FUNCTION_BLOCK FB_MotionSystem
VAR
    fbXPlanarSystem   : FB_XPlanarSystem;
    fbXPlanarMover    : ARRAY[1..maxNumMover] OF FB_XPlanarMoverStandard;
    nStartupSequence  : UDINT;
    nStartingSequence : UDINT;
    nExecutingSequence : UDINT;
    nErrorStep         : UDINT;    // step where the error happened
    nErrorID           : UDINT;    // error code of the motion command
END_VAR

METHOD Cycle
VAR
    i : UDINT;
END_VAR
// Call every PLC cycle: updates the XPlanar system and the movers.
fbXPlanarSystem.Cycle();
FOR i := 1 TO moverCount DO
    fbXPlanarMover[i].Cycle();
END_FOR
END_METHOD

METHOD Execute6DoF : BOOL
VAR_INPUT
    bReset : BOOL;
END_VAR
VAR_INST
    stStartPos   : PositionXYC;
    stCenterPos  : PositionXYC;
    stRotOptions : ST_MoveCOptions;
END_VAR
// One 6 DoF sequence with mover 1. TRUE when finished. Stops in step 900 on error.
IF bReset THEN
    Execute6DoF := FALSE;
    nExecutingSequence := 0;
    nErrorStep := 0;
    nErrorID := 0;
END_IF

CASE nExecutingSequence OF
    // store the start position
    0:  stStartPos.SetValuesXYC(fbXPlanarMover[1].P_ActPosition.x,
                                fbXPlanarMover[1].P_ActPosition.y,
                                fbXPlanarMover[1].P_ActPosition.c);
        stCenterPos.SetValuesXYC(480, 360, 0);
        stRotOptions.additionalTurns := 0;
        stRotOptions.direction := Tc3_Mc3PlanarMotion.MC_Direction.mcDirectionNonModulo;
        IF NOT bReset THEN
            nExecutingSequence := 10;
        END_IF

    // drive to the table centre
    10: fbXPlanarMover[1].MoveToPosition('To center', stCenterPos, 500, 1250, 1250, 12500);
        nExecutingSequence := 11;
    11: IF fbXPlanarMover[1].P_MoveToPosition.Done THEN
            nExecutingSequence := 20;
        ELSIF fbXPlanarMover[1].P_MoveToPosition.Error THEN
            nErrorStep := nExecutingSequence;
            nErrorID := fbXPlanarMover[1].P_MoveToPosition.ErrorID;
            nExecutingSequence := 900;
        END_IF

    // lift Z to 4 mm
    20: fbXPlanarMover[1].MoveZ('Z up', 4, 20, 100, 100, 1000);
        nExecutingSequence := 21;
    21: IF fbXPlanarMover[1].P_MoveZ.Done THEN
            nExecutingSequence := 30;
        ELSIF fbXPlanarMover[1].P_MoveZ.Error THEN
            nErrorStep := nExecutingSequence;
            nErrorID := fbXPlanarMover[1].P_MoveZ.ErrorID;
            nExecutingSequence := 900;
        END_IF

    // rotate C +90 deg
    30: fbXPlanarMover[1].MoveC('C +90', 90, 720, 1800, 1800, 9000, stRotOptions);
        nExecutingSequence := 31;
    31: IF fbXPlanarMover[1].P_MoveC.Done THEN
            nExecutingSequence := 50;
        ELSIF fbXPlanarMover[1].P_MoveC.Error THEN
            nErrorStep := nExecutingSequence;
            nErrorID := fbXPlanarMover[1].P_MoveC.ErrorID;
            nExecutingSequence := 900;
        END_IF

	// lower Z
	40: fbXPlanarMover[1].MoveZ('Z down', 2, 20, 100, 100, 1000);
        nExecutingSequence := 41;
    41: IF fbXPlanarMover[1].P_MoveZ.Done THEN
            nExecutingSequence := 100;
        ELSIF fbXPlanarMover[1].P_MoveZ.Error THEN
            nErrorStep := nExecutingSequence;
            nErrorID := fbXPlanarMover[1].P_MoveZ.ErrorID;
            nExecutingSequence := 900;
        END_IF

    // tilt A (while lifted)
    50: fbXPlanarMover[1].MoveA('A tilt', 2, 20, 100, 100, 1000);
        nExecutingSequence := 51;
    51: IF fbXPlanarMover[1].P_MoveA.Done THEN
            nExecutingSequence := 60;
        ELSIF fbXPlanarMover[1].P_MoveA.Error THEN
            nErrorStep := nExecutingSequence;
            nErrorID := fbXPlanarMover[1].P_MoveA.ErrorID;
            nExecutingSequence := 900;
        END_IF

    // tilt B
    60: fbXPlanarMover[1].MoveB('B tilt', 2, 20, 100, 100, 1000);
        nExecutingSequence := 61;
    61: IF fbXPlanarMover[1].P_MoveB.Done THEN
            nExecutingSequence := 70;
        ELSIF fbXPlanarMover[1].P_MoveB.Error THEN
            nErrorStep := nExecutingSequence;
            nErrorID := fbXPlanarMover[1].P_MoveB.ErrorID;
            nExecutingSequence := 900;
        END_IF

    // A back to 0
    70: fbXPlanarMover[1].MoveA('A back', 0, 20, 100, 100, 1000);
        nExecutingSequence := 71;
    71: IF fbXPlanarMover[1].P_MoveA.Done THEN
            nExecutingSequence := 80;
        ELSIF fbXPlanarMover[1].P_MoveA.Error THEN
            nErrorStep := nExecutingSequence;
            nErrorID := fbXPlanarMover[1].P_MoveA.ErrorID;
            nExecutingSequence := 900;
        END_IF

    // B back to 0
    80: fbXPlanarMover[1].MoveB('B back', 0, 20, 100, 100, 1000);
        nExecutingSequence := 81;
    81: IF fbXPlanarMover[1].P_MoveB.Done THEN
            nExecutingSequence := 90;
        ELSIF fbXPlanarMover[1].P_MoveB.Error THEN
            nErrorStep := nExecutingSequence;
            nErrorID := fbXPlanarMover[1].P_MoveB.ErrorID;
            nExecutingSequence := 900;
        END_IF

    // C back to 0
    90: fbXPlanarMover[1].MoveC('C back', 0, 720, 1800, 1800, 9000, stRotOptions);
        nExecutingSequence := 91;
    91: IF fbXPlanarMover[1].P_MoveC.Done THEN
            nExecutingSequence := 40;
        ELSIF fbXPlanarMover[1].P_MoveC.Error THEN
            nErrorStep := nExecutingSequence;
            nErrorID := fbXPlanarMover[1].P_MoveC.ErrorID;
            nExecutingSequence := 900;
        END_IF

    // return to the start position
    100: fbXPlanarMover[1].MoveToPosition('Back to start', stStartPos, 500, 1250, 1250, 12500);
        nExecutingSequence := 101;
    101: IF fbXPlanarMover[1].P_MoveToPosition.Done THEN
            nExecutingSequence := 110;
        ELSIF fbXPlanarMover[1].P_MoveToPosition.Error THEN
            nErrorStep := nExecutingSequence;
            nErrorID := fbXPlanarMover[1].P_MoveToPosition.ErrorID;
            nExecutingSequence := 900;
        END_IF

    // finished
    110: Execute6DoF := TRUE;

    // motion error: see nErrorStep, nErrorID
    900: ;
END_CASE
END_METHOD

METHOD Starting : BOOL
VAR_INPUT
    bReset : BOOL;
END_VAR
// Brings the system to a ready state step by step. TRUE when done.
IF bReset THEN
    Starting := FALSE;
    nStartingSequence := 0;
END_IF
CASE nStartingSequence OF
    // start
    0:  nStartingSequence := 50;
    // enable movers
    50: IF fbXPlanarSystem.EnableMovers() THEN
            nStartingSequence := 51;
        END_IF
    // wait for enable
    51: IF fbXPlanarSystem.P_EnableMovers.Done THEN
            nStartingSequence := 80;
        ELSIF fbXPlanarSystem.P_EnableMovers.Error THEN
            nStartingSequence := 90;   // enable failed
        END_IF
    // ready
    80: Starting := TRUE;
END_CASE
END_METHOD

METHOD Startup : BOOL
VAR
    i : UDINT;
END_VAR
// One-time setup: register movers (and tracks) in the system. TRUE when done.
CASE nStartupSequence OF
    0:  nStartupSequence := 1;
    1:  FOR i := 1 TO moverCount DO
            fbXPlanarSystem.SetMoverStandard(i, fbXPlanarMover[i]);
        END_FOR
        nStartupSequence := 30;
    30: Startup := TRUE;
END_CASE
END_METHOD

END_FUNCTION_BLOCK

(* stored: Version 1.1.0.1
   POU FB_MotionSystem: Id {76b90533-2f5f-4265-a888-7463c8f15552}, SpecialFunc None
   Method Cycle: Id {7a6a436f-abe3-49cf-80ba-736989644d1a}
   Method Execute6DoF: Id {8ce13323-1410-4b2b-b91c-3d53f634fa57}
   Method Starting: Id {04721e65-d0d5-4973-a78a-e55f3a27c0da}
   Method Startup: Id {ab1988d1-2b56-4e22-9706-835668cd8a23} *)
